Staubli VAL3: nmbValue.pgx

program nmbValue(num x_nStep, num x_nIndex)
  local trsf l_trsf
  local num l_nResult
begin
  switch x_nStep

    case 0
      l_trsf=savedata:fFrameItem[x_nIndex].pPointRx[0].trsf
      sUsingFrame=savedata:fFrameItem[x_nIndex].sName+" 坐标系O点"
      nNmbValue[0]=l_trsf.x
      nNmbValue[1]=l_trsf.y
      nNmbValue[2]=l_trsf.z
      nNmbValue[3]=l_trsf.rx
      nNmbValue[4]=l_trsf.ry
      nNmbValue[5]=l_trsf.rz
    break
    case 1
      l_trsf=savedata:fFrameItem[x_nIndex].pPointRx[1].trsf
      sUsingFrame=savedata:fFrameItem[x_nIndex].sName+" 坐标系X点"
      nNmbValue[0]=l_trsf.x
      nNmbValue[1]=l_trsf.y
      nNmbValue[2]=l_trsf.z
      nNmbValue[3]=l_trsf.rx
      nNmbValue[4]=l_trsf.ry
      nNmbValue[5]=l_trsf.rz
    break
    case 2
      l_trsf=savedata:fFrameItem[x_nIndex].pPointRx[2].trsf
      sUsingFrame=savedata:fFrameItem[x_nIndex].sName+" 坐标系Y点"
      nNmbValue[0]=l_trsf.x
      nNmbValue[1]=l_trsf.y
      nNmbValue[2]=l_trsf.z
      nNmbValue[3]=l_trsf.rx
      nNmbValue[4]=l_trsf.ry
      nNmbValue[5]=l_trsf.rz
    break


  endSwitch




end
